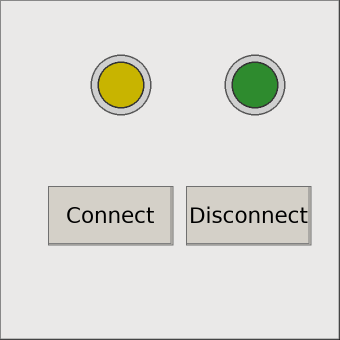
VISUALIZATION vis_FB_InterConnection  // 340x340
VAR_IN_OUT
	fb: FB_InterConnection;

END_VAR
    Rectangle (0,0 340x340)
    Button (48,186 125x59), "Connect", input disabled if: NOT fb.bAvalableToConnect
        OnMouseClick: toggle fb.reqConnect
    Button (186,186 125x59), "Disconnect", input disabled if: NOT fb.bAvalableToDisconnect
        OnMouseClick: toggle fb.reqDisconnect
    Lamp1 (220,50 70x70), variable: fb.bActive, style: Lamp-Lamp1-Green
    Lamp1 (86,50 70x70), variable: fb.bAvalableToConnect, style: Lamp-Lamp1-Yellow
END_VISUALIZATION

(* stored: Version 1.1.0.1, ProductVersion 3.1.4024.12
   Visu vis_FB_InterConnection: Id {949125f2-4032-4011-8d8a-1d74900f2da3} *)
